Fanuc KAREL source: KT00658.KL

PROGRAM KT00658
%NOLOCKGROUP
VAR
  P1: POSITION
  P2: POSITION
  OUT: INTEGER
BEGIN
  OUT = - P1
END KT00658
